(* IEC 61131-3 sources: IRIS-Project/LASAL CONTROL SOFTWARE/LasalProject_2025_09_12/Runtime/%LASALAPPDATA%/Runtime/Library/Loader/Class/MMConnectionReader, 1 file *)

(* ---- MMConnectionReader.st ---- *)
(*!
<Class
	Name               = "MMConnectionReader"
	Revision           = "0.0"
	RealtimeTask       = "false"
	CyclicTask         = "false"
	BackgroundTask     = "false"
	Sigmatek           = "true"
	OSInterface        = "false"
	HighPriority       = "false"
	Automatic          = "false"
	UpdateMode         = "Prescan"
	SharedCommandTable = "true"
	Objectsize         = "(284,120)">
	<Channels>
	</Channels>
	<RevDoku>
		<Owner Company="Sigmatek" Author="FimLuc"/>
		<Dokumentation Revision="0.0" Date="2015-10-07" Author="FimLuc" Company="Sigmatek" Description="erstell"/>
	</RevDoku>
	<Network Name="MMConnectionReader">
		<!-- List of Components in this network -->
		<Components>
			<Object
				Name       = "_base"
				Class      = "ObjectReader"
				Position   = "(218,120)"
				Visualized = "false">
				<Channels>
					<Server Name="Server0"/>
				</Channels>
			</Object>
		</Components>
		<Comments>
		</Comments>
		<!-- List of Connections in this network -->
		<Connections>
			<Connection Source="this.Server0" Destination="_base.Server0" Vertices="(690,210),(518,210),"/>
		</Connections>
		<!-- Headerfiles -->
		<Options>
		</Options>
	</Network>
</Class>
*)
#pragma using ObjectReader

MMConnectionReader : CLASS
: ObjectReader
  //Servers:
  //Clients:
  //Variables:
		pObjRd 	: ^ObjectReader;
  //Functions:

	FUNCTION GLOBAL ReadConnections
		VAR_INPUT
			pObjRd 	: ^ObjectReader;
		END_VAR;

	FUNCTION SetConn
		VAR_INPUT
			pClt 	: ^CltCh;
			iCltNr 	: UDINT;
			pThis 	: ^VirtualBase;
		END_VAR;

	FUNCTION ReadConnSmall;

	FUNCTION ReadConnLarge;
  //Tables:
	FUNCTION @STD
		VAR_OUTPUT
			ret_code	: CONFSTATES;
		END_VAR;
	FUNCTION GLOBAL TAB @CT_;
END_CLASS;

#include <RTOS_PrivHeader.h>

#pragma using MMServer

// forward declaration
FUNCTION GLOBAL _LookUpObjLex
VAR_INPUT
	pLexem     : ^CLexem;
END_VAR
VAR_OUTPUT
	ret				: ^SvrCh;
END_VAR;

(*
  liest die verbindungstabelle des on's ein
*)
FUNCTION GLOBAL MMConnectionReader::ReadConnections
	VAR_INPUT
		pObjRd 	: ^ObjectReader;
	END_VAR

  this^.pObjRd	:= pObjRd;

  ReadConnSmall();
  ReadConnLarge();

END_FUNCTION
(*
  setzt die verbindung
*)
FUNCTION MMConnectionReader::SetConn
	VAR_INPUT
		pClt 	: ^CltCh;
    iCltNr : UDINT;
    pThis	: ^VirtualBase;
	END_VAR
  VAR
    uiTry   : UINT;
    pSvr    : ^void;
    lexem   : ^CLexem;
    cCltNr : ARRAY[ 0..8 ] OF CHAR;
  END_VAR

  uiTry := pObjRd^.GetUInt();

  lexem := pObjRd^.ReadLexem();
  pSvr := _LookUpObjLex(lexem);

  IF (pSvr = NIL) THEN
       // eventuell hat das initialisieren der MMConnectionHandler zu lange gedauert,
       // sodass das MMServer-Object nocht nicht angelegt worden ist
        _itoa( iCltNr, #cCltNr[ 0 ] );
       IF(pThis <> NIL) THEN
          TRACE2_ERR("Remote object '{0}' not found. Check Stations.txt. Could not connect to object '{1}' at client {2}", #lexem^.Text[0], LSL_GetObjName(pThis), #cCltNr[ 0 ]);
       ELSE
          TRACE1_ERR("Remote object '{0}' not found. Check Stations.txt. Could not enter connection to '{1}'", #lexem^.Text[0], #cCltNr[ 0 ]);
       END_IF;
      RETURN;
  END_IF;

  IF (uiTry <> C_TRY) THEN
    pSvr$^MMServer^.m_flStatus := (pSvr$^MMServer^.m_flStatus OR MM_REQUIRED);
  END_IF;

  pClt^.pCh  := pSvr$^SvrCh;
  pClt^.pCmd := pSvr$^VirtualBase;

END_FUNCTION

FUNCTION MMConnectionReader::ReadConnSmall
VAR
  nConCnt	: UDINT;
  pClt	: ^CltCh;
  iCltNr  : UDINT;
  cCltNr : ARRAY[ 0..8 ] OF CHAR;
END_VAR

	nConCnt	:= pObjRd^.GetCount();

	IF nConCnt = 0 THEN
		RETURN;
	END_IF;

  iCltNr := 0;

	WHILE (nConCnt > 0) DO				// alle angegebenen Verbindungspaare einlesen
    iCltNr += 1;

    pClt	:= (pObjRd^.GetObjectOff()) $ ^CltCh;

    IF (pClt = NIL) THEN
      _itoa( iCltNr, #cCltNr[ 0 ] );
      TRACE0_ERR("channel '{0}' not found.", #cCltNr[ 0 ]);
			RETURN;
		END_IF;

    SetConn(pClt, iCltNr, NIL);

		nConCnt	-= 1;
	END_WHILE;

END_FUNCTION

FUNCTION MMConnectionReader::ReadConnLarge
VAR
  nConCnt	: UDINT;
  pClt	: ^CltCh;
  pThis	: ^VirtualBase;
  iCltNr  : UDINT;
  cCltNr : ARRAY[ 0..8 ] OF CHAR;
END_VAR

	nConCnt	:= pObjRd^.GetCount();

	IF nConCnt = 0 THEN
		RETURN;
	END_IF;

  iCltNr := 0;

	WHILE (nConCnt > 0) DO				// alle angegebenen Verbindungspaare einlesen
    iCltNr += 1;
		pThis	:= pObjRd^.GetObjectNo();
		pClt	:= pObjRd^.GetChPtr(pThis);
    IF (pClt = NIL) THEN
      _itoa( iCltNr, #cCltNr[ 0 ] );
      TRACE1_ERR("Channel '{0}' of Object '{1}' not found.", #cCltNr[ 0 ], LSL_GetObjName(pThis));
			RETURN;
		END_IF;

    SetConn(pClt, iCltNr, pThis);

		nConCnt	-= 1;
	END_WHILE;

END_FUNCTION
